Fanuc KAREL source: KT00768.KL

PROGRAM KT00768
%NOLOCKGROUP
VAR
  B1: BOOLEAN
  B2: BOOLEAN
  OUT: INTEGER
BEGIN
  B1 = TRUE
  B2 = FALSE
  B1 = TRUE
  B2 = FALSE
  OUT = ACOS(B1)
END KT00768
